INTERFACE I_MoverDisableAlgorithm EXTENDS i_Task


METHOD Abort : HRESULT
VAR_INPUT
END_VAR
END_METHOD

METHOD Disable : HRESULT
VAR_INPUT
END_VAR
END_METHOD

METHOD Reset : HRESULT
VAR_INPUT
END_VAR
END_METHOD

METHOD SetComponents : BOOL
VAR_INPUT
	MoverArray : ARRAY[0..TcIoXtsEnvironmentParameterList.MaxXtsMoversPerXpu] OF I_XtsMover;
	CAGroup : I_CollisionGroup;
	MoverCount : UDINT;
END_VAR
END_METHOD

END_INTERFACE

(* stored: Version 1.1.0.1
   Itf I_MoverDisableAlgorithm: Id {88d2d5be-93c8-4054-ba32-89a88adb2d09}
   Method Abort: Id {ca15dffc-ad96-49a0-8b36-c8b86b1ddeee}
   Method Disable: Id {bc955e12-7352-42fe-b966-d4b86508eddb}
   Method Reset: Id {2f514183-d44a-4af8-bf34-d4b92afcf649}
   Method SetComponents: Id {02927f80-cee4-4ccc-bf30-7be3bd61e23c} *)
